(* IEC 61131-3 sources: trust-platform/tests/fixtures/hmi_reliability_bundle/sources, 2 files *)

(* ---- config.st ---- *)
CONFIGURATION Config
VAR_GLOBAL
    InSignal AT %IX0.0 : BOOL;
    OutSignal AT %QX0.0 : BOOL;
END_VAR

RESOURCE ReliabilityResource ON PLC
    TASK MainTask (INTERVAL := T#100ms, PRIORITY := 1);
    PROGRAM P1 WITH MainTask : Main;
END_RESOURCE
END_CONFIGURATION

(* ---- main.st ---- *)
PROGRAM Main
VAR
    Count : INT := 0;
END_VAR

VAR_EXTERNAL
    InSignal : BOOL;
    OutSignal : BOOL;
END_VAR

IF InSignal THEN
    Count := Count + 1;
END_IF;

OutSignal := (Count MOD 2) = 1;
END_PROGRAM
